PROGRAM main
  VAR
    B1 AT %IX0.0     : BOOL; (* sensor de cajas *)
    KM1 AT %QX0.0    : BOOL; (* banda (bobina 00001 para la PC) *)
    CAJAS AT %MW0    : INT; (* holding 40001: cajas contadas *)
    P_MARCHA AT %MW1 : INT; (* holding 40002: pulsador remoto MARCHA *)
    P_PARO AT %MW2   : INT; (* holding 40003: pulsador remoto PARO *)
    P_CERO AT %MW3   : INT; (* holding 40004: pulsador remoto contador a cero *)
    F_CAJA           : R_TRIG;
    O_MARCHA         : BOOL; (* la PC pidió marcha *)
    O_PARO           : BOOL; (* la PC pidió paro *)
    O_CERO           : BOOL; (* la PC pidió el contador a cero *)
  END_VAR
  VAR  (* added by the conversion: wires and edge detectors of the diagram *)
    R_TRIG1 : R_TRIG;
  END_VAR

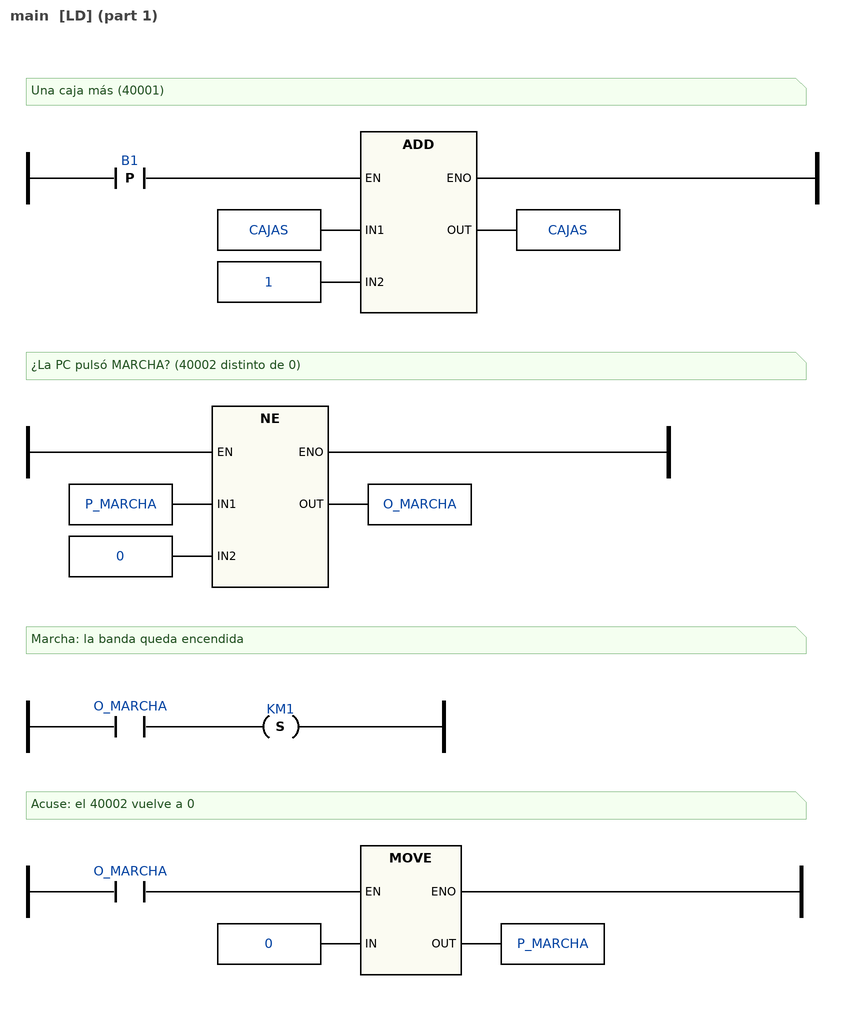
(* LD diagram, written out as Structured Text *)
(* Una caja más (40001) *)
R_TRIG1(CLK := B1);
IF R_TRIG1.Q THEN CAJAS := CAJAS + 1; END_IF;
(* ¿La PC pulsó MARCHA? (40002 distinto de 0) *)
O_MARCHA := P_MARCHA <> 0;
(* Marcha: la banda queda encendida *)
IF O_MARCHA THEN KM1 := TRUE; END_IF;
(* Acuse: el 40002 vuelve a 0 *)
IF O_MARCHA THEN P_MARCHA := 0; END_IF;
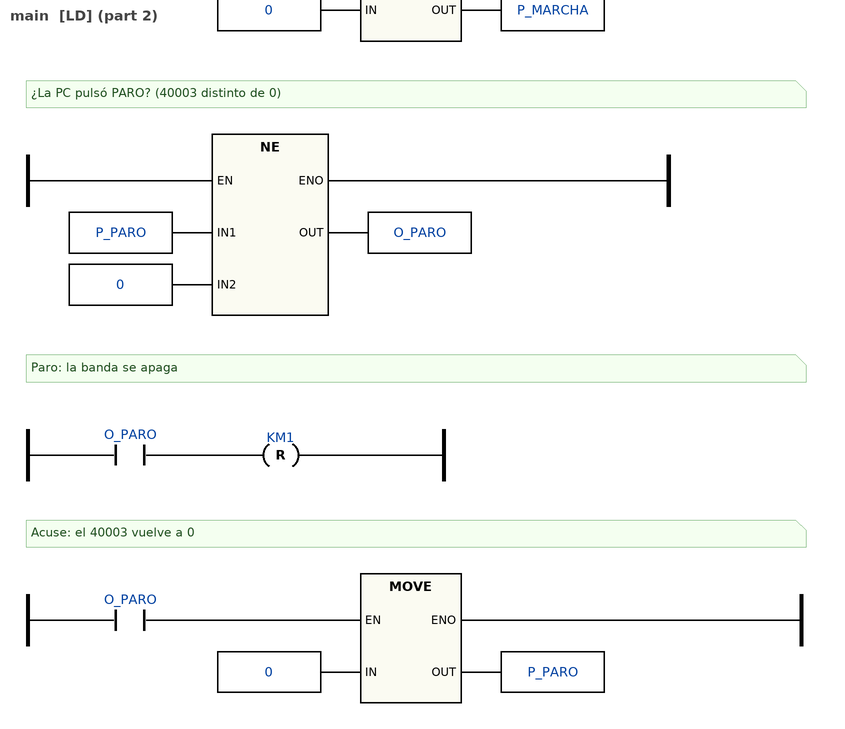
(* ¿La PC pulsó PARO? (40003 distinto de 0) *)
O_PARO := P_PARO <> 0;
(* Paro: la banda se apaga *)
IF O_PARO THEN KM1 := FALSE; END_IF;
(* Acuse: el 40003 vuelve a 0 *)
IF O_PARO THEN P_PARO := 0; END_IF;
END_PROGRAM
